(* IEC 61131-3 sources: PortalRobot/Portal_robot/Device/application/ST/ST_TEST, 4 files *)

(* ---- E_CELL_TEST_ENVIRONMENT.st ---- *)
{attribute 'qualified_only'}
TYPE E_CELL_TEST_ENVIRONMENT :
(
	NORMAL := 0,
	SIMULATION := 1,
	SC500_BENCH := 2
);
END_TYPE

(* ---- E_TEST_SPEED_PROFILE.st ---- *)
{attribute 'qualified_only'}
TYPE E_TEST_SPEED_PROFILE :
(
	REALTIME := 0,
	FAST := 1
);
END_TYPE

(* ---- ST_TEST_OBSERVABILITY.st ---- *)
TYPE ST_TEST_OBSERVABILITY :
STRUCT
	udiAppliedScenarioSeq : UDINT;
	uiSchemaVersion : UINT;
	uiReturnMagazine : UINT;
	uiCellState : UINT;
	uiRobotState : UINT;
	uiRobotAction : UINT;
	uiRobotPoint : UINT;
	uiActiveMagazine : UINT;
	uiMagazineState : UINT;
	uiMagazineOperation : UINT;
	uiTakeSlot : UINT;
	uiPutSlot : UINT;
	auiMachineState : ARRAY [1..3] OF UINT;
	auiMachineOperation : ARRAY [1..3] OF UINT;
	uiSelectedMachine : UINT;
	uiSelectedType : UINT;
	uiErrorSource : UINT;
	dwErrorCode : DWORD;
END_STRUCT
END_TYPE

(* ---- ST_TEST_SCENARIO_BUFFER.st ---- *)
TYPE ST_TEST_SCENARIO_BUFFER :
STRUCT
	udiLoadSeq : UDINT;
	uiSchemaVersion : UINT; // v3: explicit magazine owner and both pallets
	uiMagazineMode : UINT; // Must match the selected mode; never switches mechanics
	axOperatorLoaded : ARRAY [1..2] OF BOOL;
	axAutoSwap : ARRAY [1..2] OF BOOL;
	aauiOperatorSlotContent : ARRAY [1..2, 1..120] OF UINT; // 1..96 in twin mode
	axGeometryEnabled : ARRAY [1..2] OF BOOL;
	axGeometryCall : ARRAY [1..3] OF BOOL;
	xGeometryWaitWhenOccupied : BOOL;
	uiTypeCount : UINT;
	axMagazineEnabled : ARRAY [1..2] OF BOOL;
	auiMachineState : ARRAY [1..3] OF UINT; // 0 disabled, 1 empty, 2 blank processing, 3 detail ready
	auiMachineType : ARRAY [1..3] OF UINT;
	aauiSlotContent : ARRAY [1..2, 1..120] OF UINT; // Robot-side slots: static 1..120; twin 1..96; 0 empty, 1 blank, 2 detail
	auiSlotType : ARRAY [1..120] OF UINT;
	auiGripperContent : ARRAY [1..2] OF UINT;
	auiGripperType : ARRAY [1..2] OF UINT;
	uiOrientation : UINT; // 0 blank, 1 detail
	dwCellFaultMask : DWORD; // b0: противоречивое наличие детали в обоих захватах
	dwRobotFaultMask : DWORD; // b0 wrong action; b1..b4 grippers; b5..b8 point validation
	adwMagazineFaultMask : ARRAY [1..2] OF DWORD; // b0 wrong op; b1 no blank; b2 no slot; b3 invalid slot; b4 content; b5 geometry
	adwMachineFaultMask : ARRAY [1..3] OF DWORD; // b0 alarm; b1 door; b2 chuck; b3..b10 timeouts
END_STRUCT
END_TYPE
